(* IEC 61131-3 sources: PLC-Static-Analysis/modules/plc-rules/src/test/resources/PLCA-Q008/library, 1 file *)

(* ---- lib.st ---- *)
FUNCTION F_Scale : REAL
VAR_INPUT
    r : REAL;
END_VAR
F_Scale := r * 2.0;
END_FUNCTION

FUNCTION_BLOCK FB_Filter
VAR
    r : REAL;
END_VAR
r := r * 0.5;
END_FUNCTION_BLOCK
